// TIA Portal V20 export
// export: Created 2026-10-19T18:07:47.4459135Z, ExportSetting None, DisplayName Totally Integrated Automation Portal, DisplayVersion V20 Update 6, DisplayName TIA Portal Openness, DisplayVersion V20 Update 6, DisplayName TIA Portal Version Control Interface, DisplayVersion V20 Update 6, DisplayName SINAMICS Startdrive Advanced, DisplayVersion V20 SP1, DisplayName SINAMICS Startdrive G130, G150, S120, S150, SINAMICS MV, G220, S200, S210, DisplayVersion V20 SP1, DisplayName SINAMICS Startdrive G110M, G120, G120C, G120D, G120P, G115D, DisplayVersion V20 SP1, DisplayName STEP 7 Professional, DisplayVersion V20 Update 6, DisplayName STEP 7 Safety, DisplayVersion V20 Update 2, DisplayName WinCC Basic/Comfort/Advanced, DisplayVersion V20 Update 6, DisplayName WinCC Unified, DisplayVersion V20 Update 6
VAR_GLOBAL   // PLC tag table "Errors"
   Errors_IND360_Smart5_Red_Level_5 AT %MW700 : Word;
   Error AT %M729.0 : Bool;
   Errors_Profinet_1 AT %MW730 : Word;
   Errors_Profinet_2 AT %MW732 : Word;
   Errors_Profinet_3 AT %MW734 : Word;
   Erros_LMs_1 AT %MW736 : Word;
   Erros_LMs_2 AT %MW738 : Word;
   Erros_LMs_3 AT %MW740 : Word;
   "IND_360_SB Status Group 1" AT %MW742 : Word;
   Error_Devices AT %MW744 : Word;
   "Sick Lector_Error code 1" AT %MW746 : Word;
   "Sick Lector_Error code 2" AT %MW748 : Word;
   "Linear Encoder_Device Errors" AT %MW750 : Word;
   "Linear Encoder_Warnings" AT %MW752 : Word;
END_VAR
